DATA_BLOCK "LatchInstance"
{ S7_Optimized_Access := 'TRUE' }
VERSION : 0.1
"FB_BasicLatch"
BEGIN
END_DATA_BLOCK
